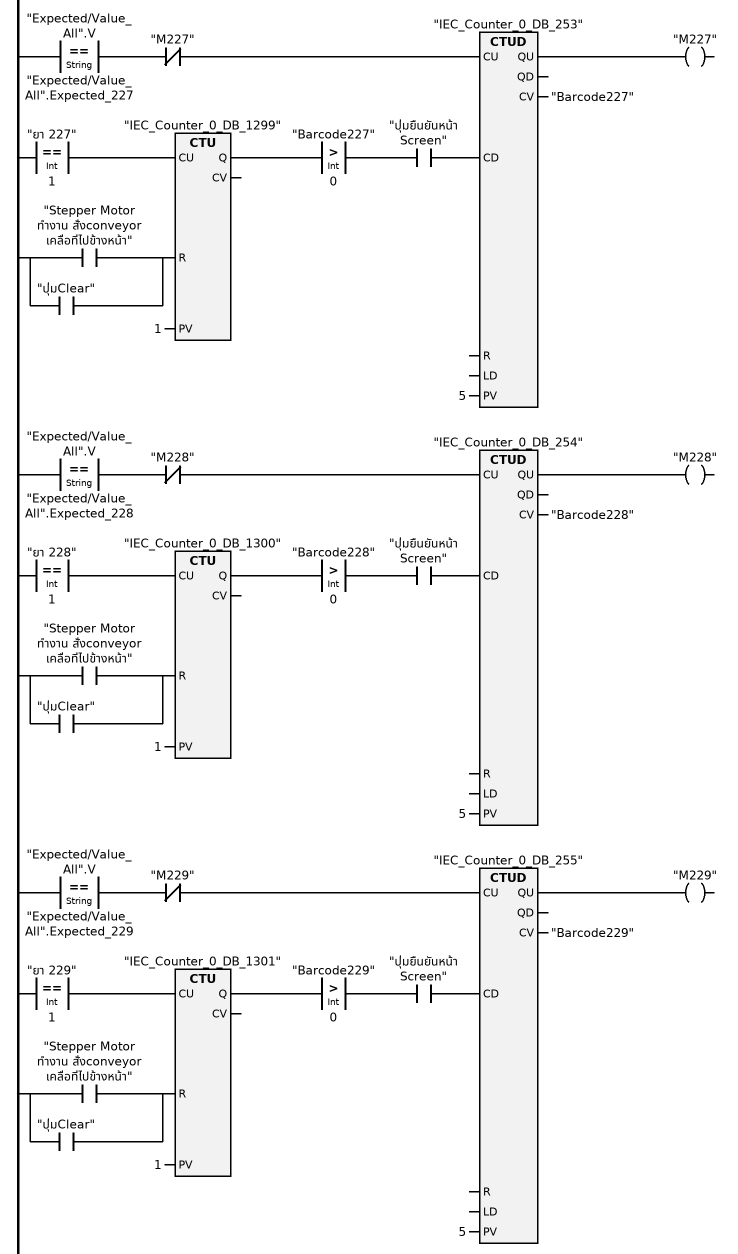
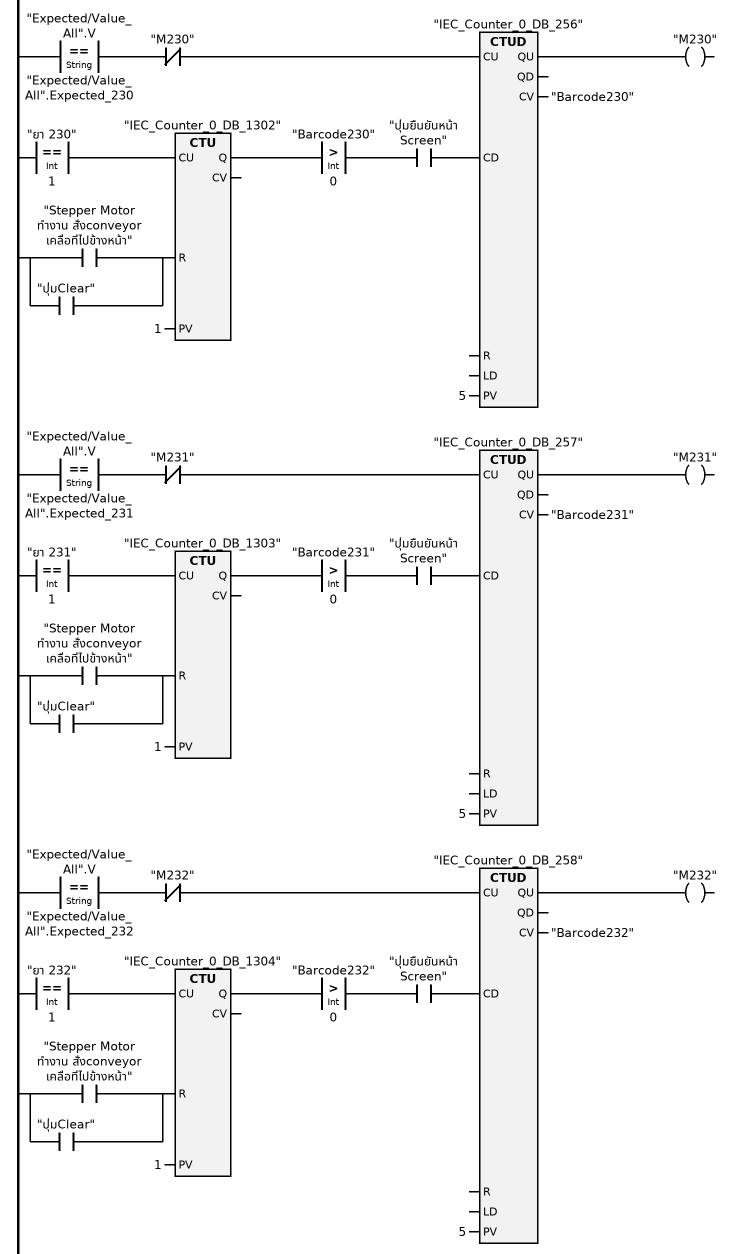
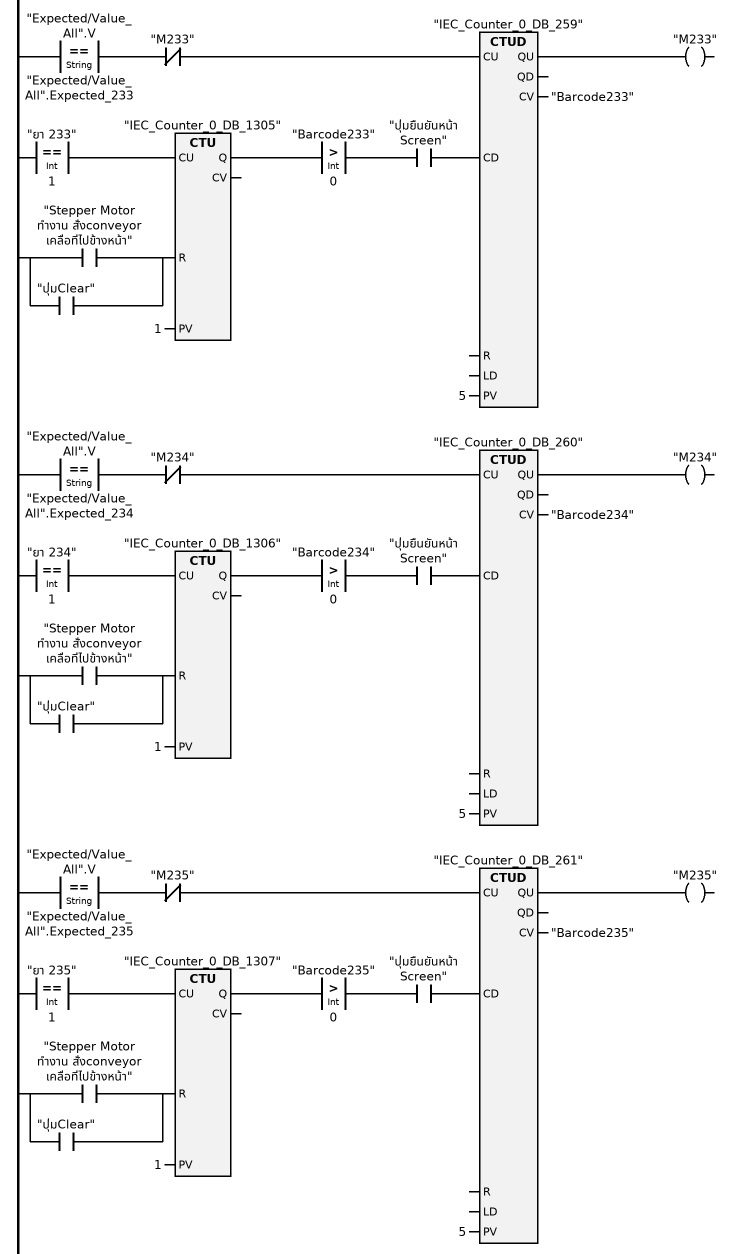
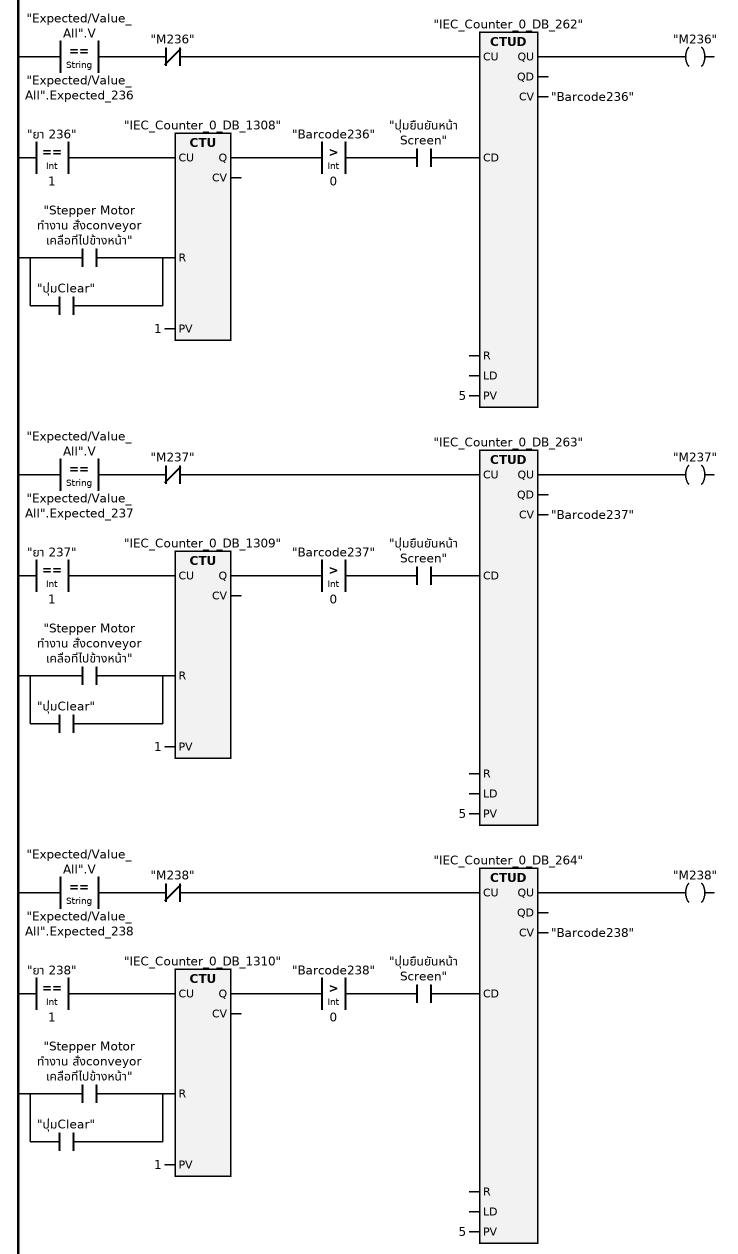
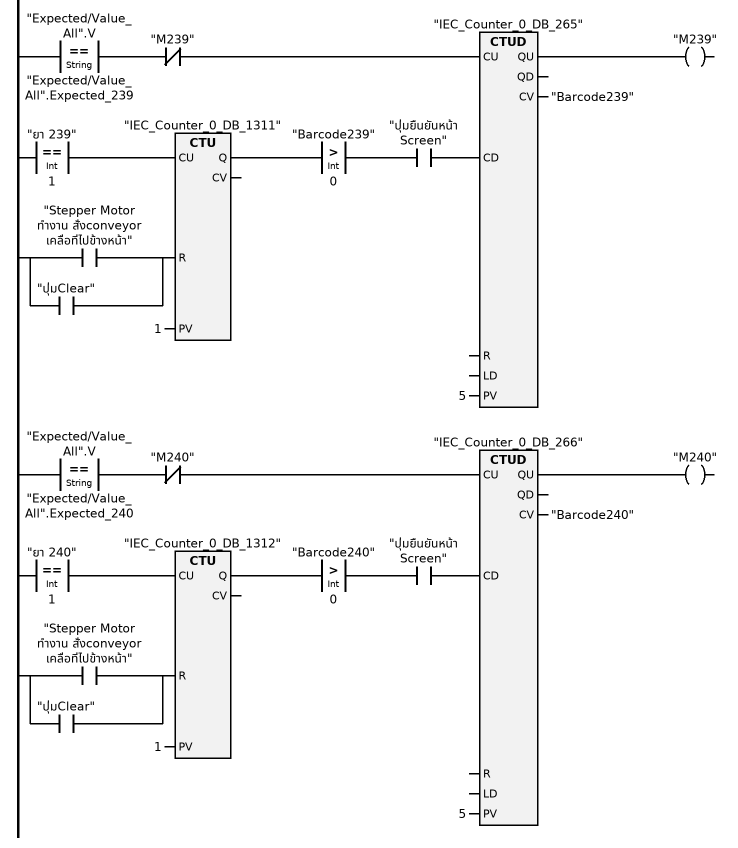
   "IEC_Counter_0_DB_1293".CTU(CU := "ยา 221" = 1,
                           R := "Stepper Motor ทำงาน สั่งconveyor เคลื่อที่ไปข้างหน้า" OR "ปุ่มClear",
                           PV := 1);
   "IEC_Counter_0_DB_247".CTUD(CU := ("Expected/Value_All".V = "Expected/Value_All".Expected_221) AND NOT "M221",
                           CD := "IEC_Counter_0_DB_1293".Q AND ("Barcode221" > 0) AND "ปุ่มยืนยันหน้า Screen",
                           PV := 5,
                           CV => "Barcode221");
   "M221" := "IEC_Counter_0_DB_247".QU;
   "IEC_Counter_0_DB_1294".CTU(CU := "ยา 222" = 1,
                           R := "Stepper Motor ทำงาน สั่งconveyor เคลื่อที่ไปข้างหน้า" OR "ปุ่มClear",
                           PV := 1);
   "IEC_Counter_0_DB_248".CTUD(CU := ("Expected/Value_All".V = "Expected/Value_All".Expected_222) AND NOT "M222",
                           CD := "IEC_Counter_0_DB_1294".Q AND ("Barcode222" > 0) AND "ปุ่มยืนยันหน้า Screen",
                           PV := 5,
                           CV => "Barcode222");
   "M222" := "IEC_Counter_0_DB_248".QU;
   "IEC_Counter_0_DB_1295".CTU(CU := "ยา 223" = 1,
                           R := "Stepper Motor ทำงาน สั่งconveyor เคลื่อที่ไปข้างหน้า" OR "ปุ่มClear",
                           PV := 1);
   "IEC_Counter_0_DB_249".CTUD(CU := ("Expected/Value_All".V = "Expected/Value_All".Expected_223) AND NOT "M223",
                           CD := "IEC_Counter_0_DB_1295".Q AND ("Barcode223" > 0) AND "ปุ่มยืนยันหน้า Screen",
                           PV := 5,
                           CV => "Barcode223");
   "M223" := "IEC_Counter_0_DB_249".QU;
   "IEC_Counter_0_DB_1296".CTU(CU := "ยา 224" = 1,
                           R := "Stepper Motor ทำงาน สั่งconveyor เคลื่อที่ไปข้างหน้า" OR "ปุ่มClear",
                           PV := 1);
   "IEC_Counter_0_DB_250".CTUD(CU := ("Expected/Value_All".V = "Expected/Value_All".Expected_224) AND NOT "M224",
                           CD := "IEC_Counter_0_DB_1296".Q AND ("Barcode224" > 0) AND "ปุ่มยืนยันหน้า Screen",
                           PV := 5,
                           CV => "Barcode224");
   "M224" := "IEC_Counter_0_DB_250".QU;
   "IEC_Counter_0_DB_1297".CTU(CU := "ยา 225" = 1,
                           R := "Stepper Motor ทำงาน สั่งconveyor เคลื่อที่ไปข้างหน้า" OR "ปุ่มClear",
                           PV := 1);
   "IEC_Counter_0_DB_251".CTUD(CU := ("Expected/Value_All".V = "Expected/Value_All".Expected_225) AND NOT "M225",
                           CD := "IEC_Counter_0_DB_1297".Q AND ("Barcode225" > 0) AND "ปุ่มยืนยันหน้า Screen",
                           PV := 5,
                           CV => "Barcode225");
   "M225" := "IEC_Counter_0_DB_251".QU;
   "IEC_Counter_0_DB_1298".CTU(CU := "ยา 226" = 1,
                           R := "Stepper Motor ทำงาน สั่งconveyor เคลื่อที่ไปข้างหน้า" OR "ปุ่มClear",
                           PV := 1);
   "IEC_Counter_0_DB_252".CTUD(CU := ("Expected/Value_All".V = "Expected/Value_All".Expected_226) AND NOT "M226",
                           CD := "IEC_Counter_0_DB_1298".Q AND ("Barcode226" > 0) AND "ปุ่มยืนยันหน้า Screen",
                           PV := 5,
                           CV => "Barcode226");
   "M226" := "IEC_Counter_0_DB_252".QU;
   "IEC_Counter_0_DB_1299".CTU(CU := "ยา 227" = 1,
                           R := "Stepper Motor ทำงาน สั่งconveyor เคลื่อที่ไปข้างหน้า" OR "ปุ่มClear",
                           PV := 1);
   "IEC_Counter_0_DB_253".CTUD(CU := ("Expected/Value_All".V = "Expected/Value_All".Expected_227) AND NOT "M227",
                           CD := "IEC_Counter_0_DB_1299".Q AND ("Barcode227" > 0) AND "ปุ่มยืนยันหน้า Screen",
                           PV := 5,
                           CV => "Barcode227");
   "M227" := "IEC_Counter_0_DB_253".QU;
   "IEC_Counter_0_DB_1300".CTU(CU := "ยา 228" = 1,
                           R := "Stepper Motor ทำงาน สั่งconveyor เคลื่อที่ไปข้างหน้า" OR "ปุ่มClear",
                           PV := 1);
   "IEC_Counter_0_DB_254".CTUD(CU := ("Expected/Value_All".V = "Expected/Value_All".Expected_228) AND NOT "M228",
                           CD := "IEC_Counter_0_DB_1300".Q AND ("Barcode228" > 0) AND "ปุ่มยืนยันหน้า Screen",
                           PV := 5,
                           CV => "Barcode228");
   "M228" := "IEC_Counter_0_DB_254".QU;
   "IEC_Counter_0_DB_1301".CTU(CU := "ยา 229" = 1,
                           R := "Stepper Motor ทำงาน สั่งconveyor เคลื่อที่ไปข้างหน้า" OR "ปุ่มClear",
                           PV := 1);
   "IEC_Counter_0_DB_255".CTUD(CU := ("Expected/Value_All".V = "Expected/Value_All".Expected_229) AND NOT "M229",
                           CD := "IEC_Counter_0_DB_1301".Q AND ("Barcode229" > 0) AND "ปุ่มยืนยันหน้า Screen",
                           PV := 5,
                           CV => "Barcode229");
   "M229" := "IEC_Counter_0_DB_255".QU;
   "IEC_Counter_0_DB_1302".CTU(CU := "ยา 230" = 1,
                           R := "Stepper Motor ทำงาน สั่งconveyor เคลื่อที่ไปข้างหน้า" OR "ปุ่มClear",
                           PV := 1);
   "IEC_Counter_0_DB_256".CTUD(CU := ("Expected/Value_All".V = "Expected/Value_All".Expected_230) AND NOT "M230",
                           CD := "IEC_Counter_0_DB_1302".Q AND ("Barcode230" > 0) AND "ปุ่มยืนยันหน้า Screen",
                           PV := 5,
                           CV => "Barcode230");
   "M230" := "IEC_Counter_0_DB_256".QU;
   "IEC_Counter_0_DB_1303".CTU(CU := "ยา 231" = 1,
                           R := "Stepper Motor ทำงาน สั่งconveyor เคลื่อที่ไปข้างหน้า" OR "ปุ่มClear",
                           PV := 1);
   "IEC_Counter_0_DB_257".CTUD(CU := ("Expected/Value_All".V = "Expected/Value_All".Expected_231) AND NOT "M231",
                           CD := "IEC_Counter_0_DB_1303".Q AND ("Barcode231" > 0) AND "ปุ่มยืนยันหน้า Screen",
                           PV := 5,
                           CV => "Barcode231");
   "M231" := "IEC_Counter_0_DB_257".QU;
   "IEC_Counter_0_DB_1304".CTU(CU := "ยา 232" = 1,
                           R := "Stepper Motor ทำงาน สั่งconveyor เคลื่อที่ไปข้างหน้า" OR "ปุ่มClear",
                           PV := 1);
   "IEC_Counter_0_DB_258".CTUD(CU := ("Expected/Value_All".V = "Expected/Value_All".Expected_232) AND NOT "M232",
                           CD := "IEC_Counter_0_DB_1304".Q AND ("Barcode232" > 0) AND "ปุ่มยืนยันหน้า Screen",
                           PV := 5,
                           CV => "Barcode232");
   "M232" := "IEC_Counter_0_DB_258".QU;
   "IEC_Counter_0_DB_1305".CTU(CU := "ยา 233" = 1,
                           R := "Stepper Motor ทำงาน สั่งconveyor เคลื่อที่ไปข้างหน้า" OR "ปุ่มClear",
                           PV := 1);
   "IEC_Counter_0_DB_259".CTUD(CU := ("Expected/Value_All".V = "Expected/Value_All".Expected_233) AND NOT "M233",
                           CD := "IEC_Counter_0_DB_1305".Q AND ("Barcode233" > 0) AND "ปุ่มยืนยันหน้า Screen",
                           PV := 5,
                           CV => "Barcode233");
   "M233" := "IEC_Counter_0_DB_259".QU;
   "IEC_Counter_0_DB_1306".CTU(CU := "ยา 234" = 1,
                           R := "Stepper Motor ทำงาน สั่งconveyor เคลื่อที่ไปข้างหน้า" OR "ปุ่มClear",
                           PV := 1);
   "IEC_Counter_0_DB_260".CTUD(CU := ("Expected/Value_All".V = "Expected/Value_All".Expected_234) AND NOT "M234",
                           CD := "IEC_Counter_0_DB_1306".Q AND ("Barcode234" > 0) AND "ปุ่มยืนยันหน้า Screen",
                           PV := 5,
                           CV => "Barcode234");
   "M234" := "IEC_Counter_0_DB_260".QU;
   "IEC_Counter_0_DB_1307".CTU(CU := "ยา 235" = 1,
                           R := "Stepper Motor ทำงาน สั่งconveyor เคลื่อที่ไปข้างหน้า" OR "ปุ่มClear",
                           PV := 1);
   "IEC_Counter_0_DB_261".CTUD(CU := ("Expected/Value_All".V = "Expected/Value_All".Expected_235) AND NOT "M235",
                           CD := "IEC_Counter_0_DB_1307".Q AND ("Barcode235" > 0) AND "ปุ่มยืนยันหน้า Screen",
                           PV := 5,
                           CV => "Barcode235");
   "M235" := "IEC_Counter_0_DB_261".QU;
   "IEC_Counter_0_DB_1308".CTU(CU := "ยา 236" = 1,
                           R := "Stepper Motor ทำงาน สั่งconveyor เคลื่อที่ไปข้างหน้า" OR "ปุ่มClear",
                           PV := 1);
   "IEC_Counter_0_DB_262".CTUD(CU := ("Expected/Value_All".V = "Expected/Value_All".Expected_236) AND NOT "M236",
                           CD := "IEC_Counter_0_DB_1308".Q AND ("Barcode236" > 0) AND "ปุ่มยืนยันหน้า Screen",
                           PV := 5,
                           CV => "Barcode236");
   "M236" := "IEC_Counter_0_DB_262".QU;
   "IEC_Counter_0_DB_1309".CTU(CU := "ยา 237" = 1,
                           R := "Stepper Motor ทำงาน สั่งconveyor เคลื่อที่ไปข้างหน้า" OR "ปุ่มClear",
                           PV := 1);
   "IEC_Counter_0_DB_263".CTUD(CU := ("Expected/Value_All".V = "Expected/Value_All".Expected_237) AND NOT "M237",
                           CD := "IEC_Counter_0_DB_1309".Q AND ("Barcode237" > 0) AND "ปุ่มยืนยันหน้า Screen",
                           PV := 5,
                           CV => "Barcode237");
   "M237" := "IEC_Counter_0_DB_263".QU;
   "IEC_Counter_0_DB_1310".CTU(CU := "ยา 238" = 1,
                           R := "Stepper Motor ทำงาน สั่งconveyor เคลื่อที่ไปข้างหน้า" OR "ปุ่มClear",
                           PV := 1);
   "IEC_Counter_0_DB_264".CTUD(CU := ("Expected/Value_All".V = "Expected/Value_All".Expected_238) AND NOT "M238",
                           CD := "IEC_Counter_0_DB_1310".Q AND ("Barcode238" > 0) AND "ปุ่มยืนยันหน้า Screen",
                           PV := 5,
                           CV => "Barcode238");
   "M238" := "IEC_Counter_0_DB_264".QU;
   "IEC_Counter_0_DB_1311".CTU(CU := "ยา 239" = 1,
                           R := "Stepper Motor ทำงาน สั่งconveyor เคลื่อที่ไปข้างหน้า" OR "ปุ่มClear",
                           PV := 1);
   "IEC_Counter_0_DB_265".CTUD(CU := ("Expected/Value_All".V = "Expected/Value_All".Expected_239) AND NOT "M239",
                           CD := "IEC_Counter_0_DB_1311".Q AND ("Barcode239" > 0) AND "ปุ่มยืนยันหน้า Screen",
                           PV := 5,
                           CV => "Barcode239");
   "M239" := "IEC_Counter_0_DB_265".QU;
   "IEC_Counter_0_DB_1312".CTU(CU := "ยา 240" = 1,
                           R := "Stepper Motor ทำงาน สั่งconveyor เคลื่อที่ไปข้างหน้า" OR "ปุ่มClear",
                           PV := 1);
   "IEC_Counter_0_DB_266".CTUD(CU := ("Expected/Value_All".V = "Expected/Value_All".Expected_240) AND NOT "M240",
                           CD := "IEC_Counter_0_DB_1312".Q AND ("Barcode240" > 0) AND "ปุ่มยืนยันหน้า Screen",
                           PV := 5,
                           CV => "Barcode240");
   "M240" := "IEC_Counter_0_DB_266".QU;
END_REGION

REGION Network 13
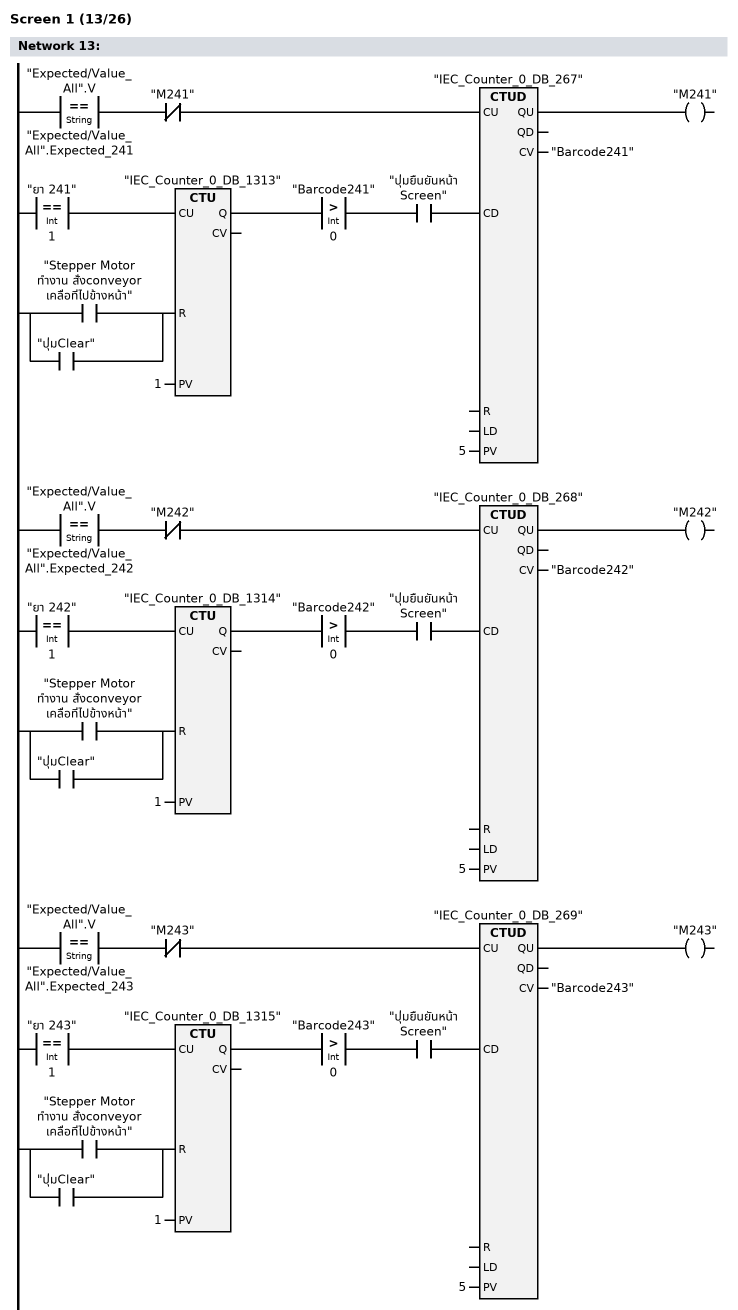
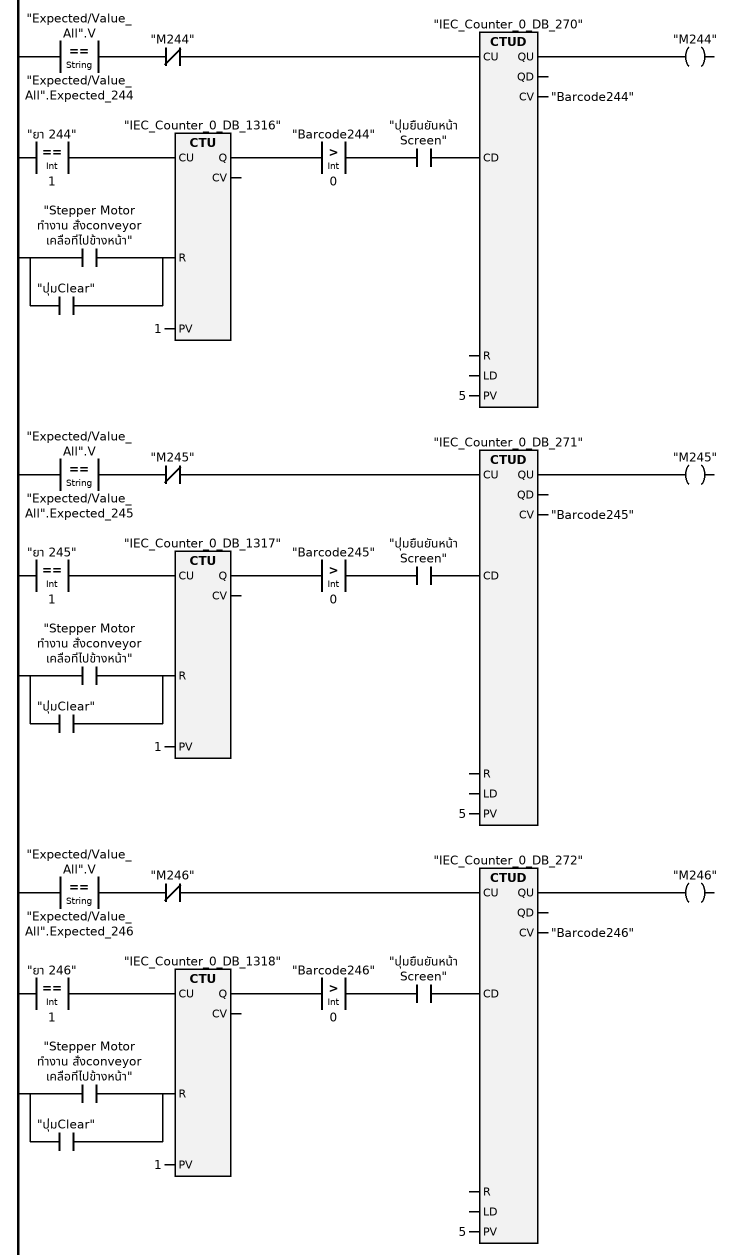
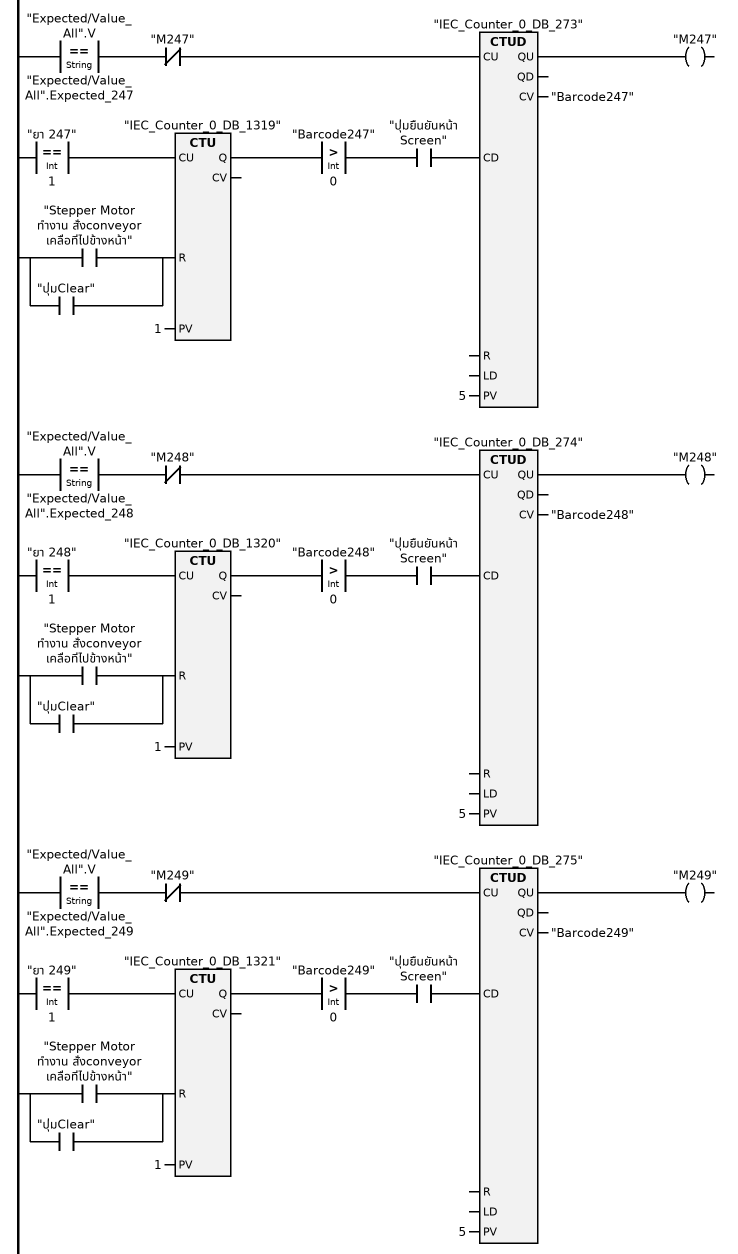
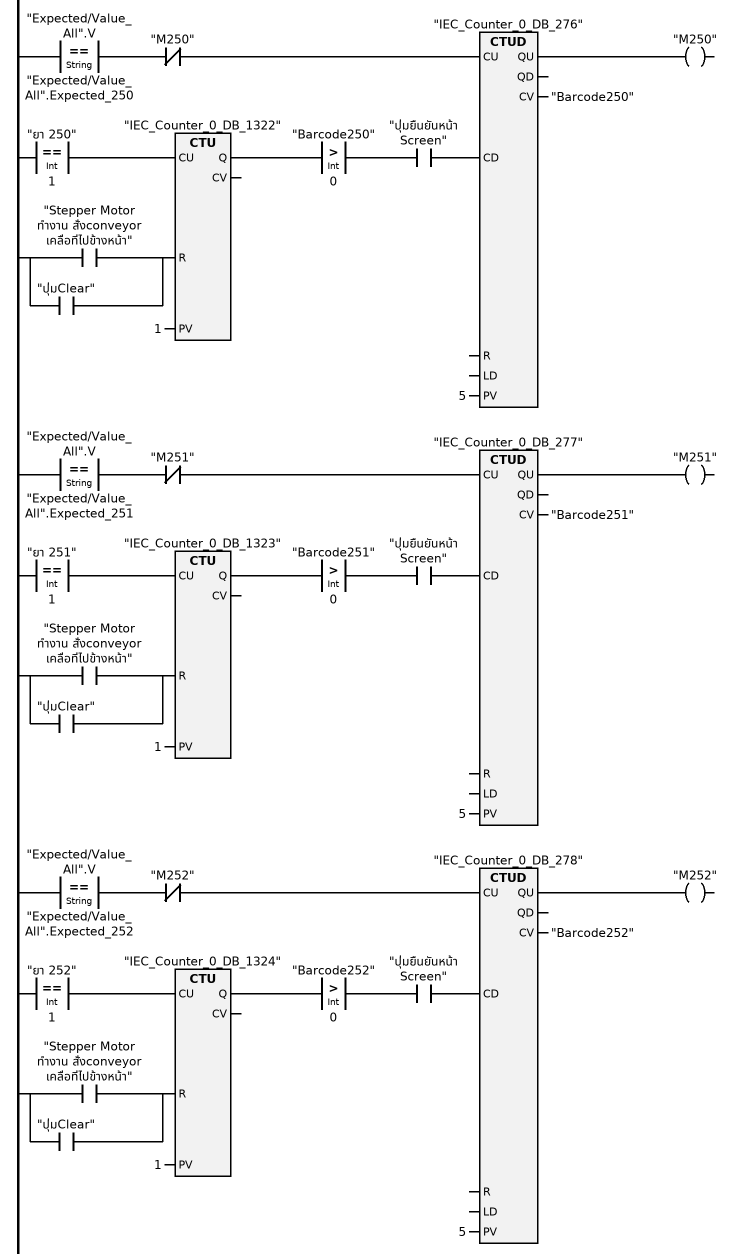
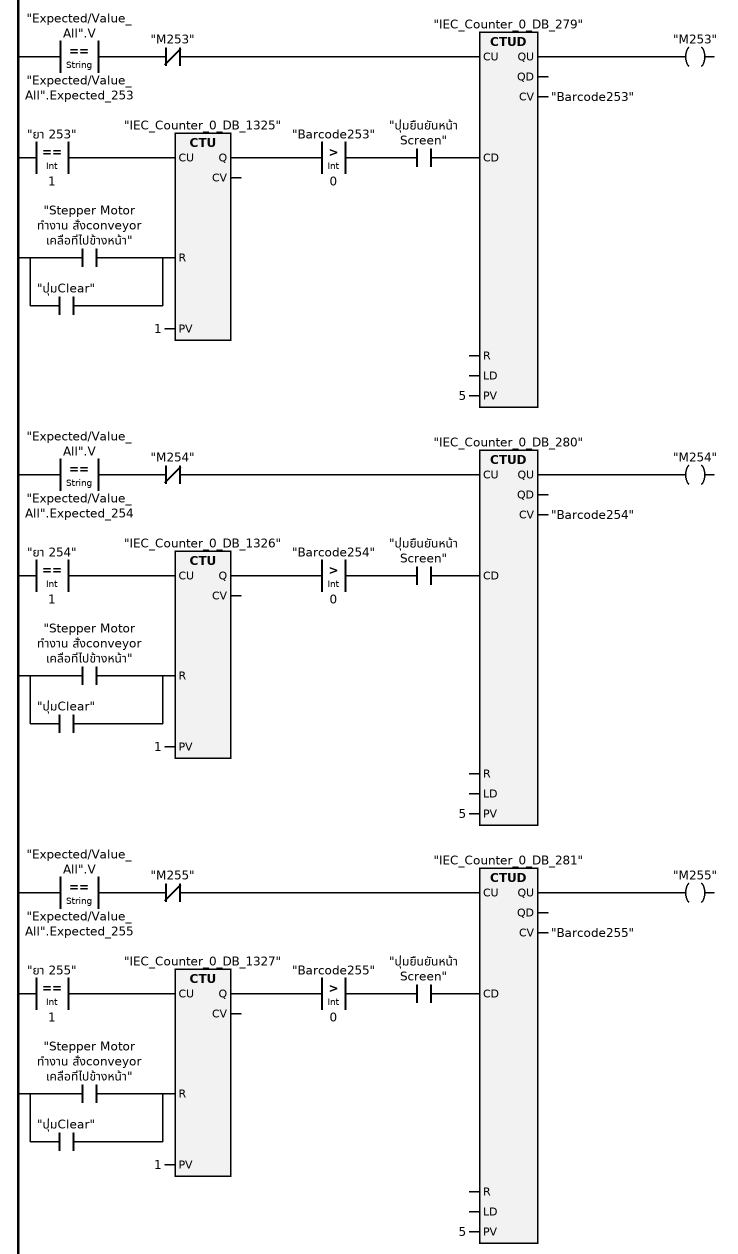
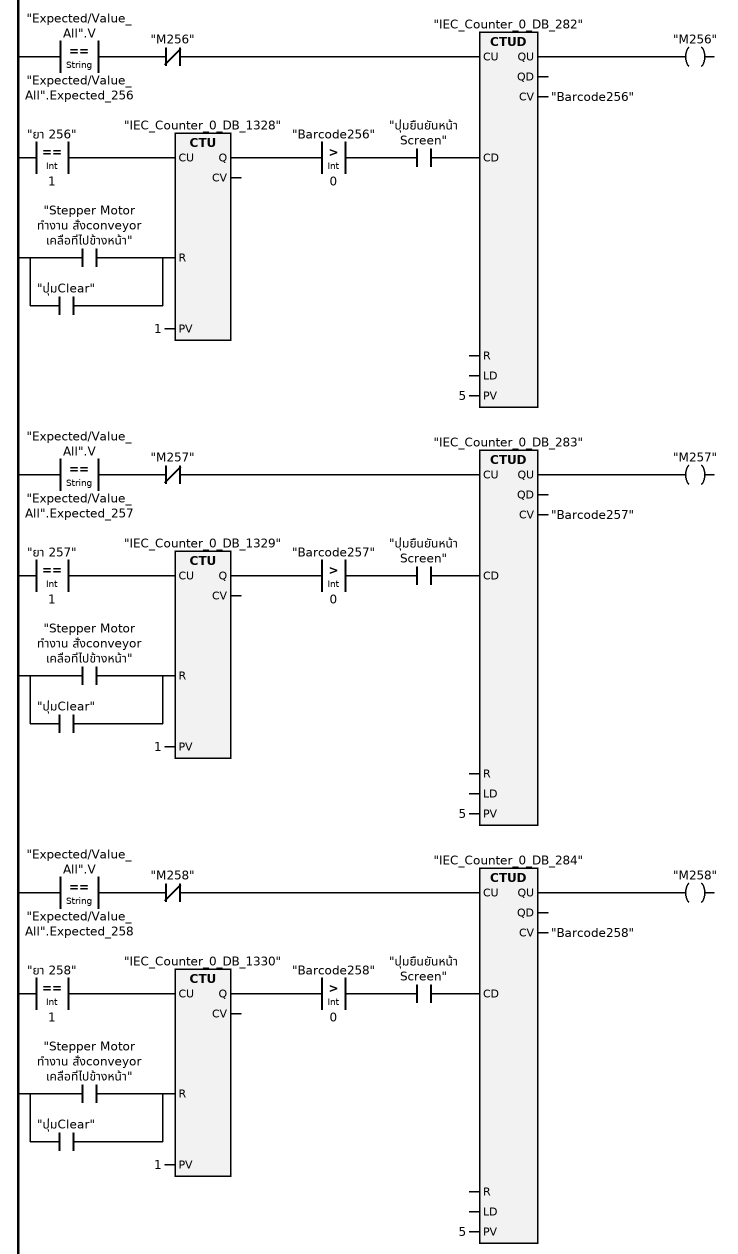
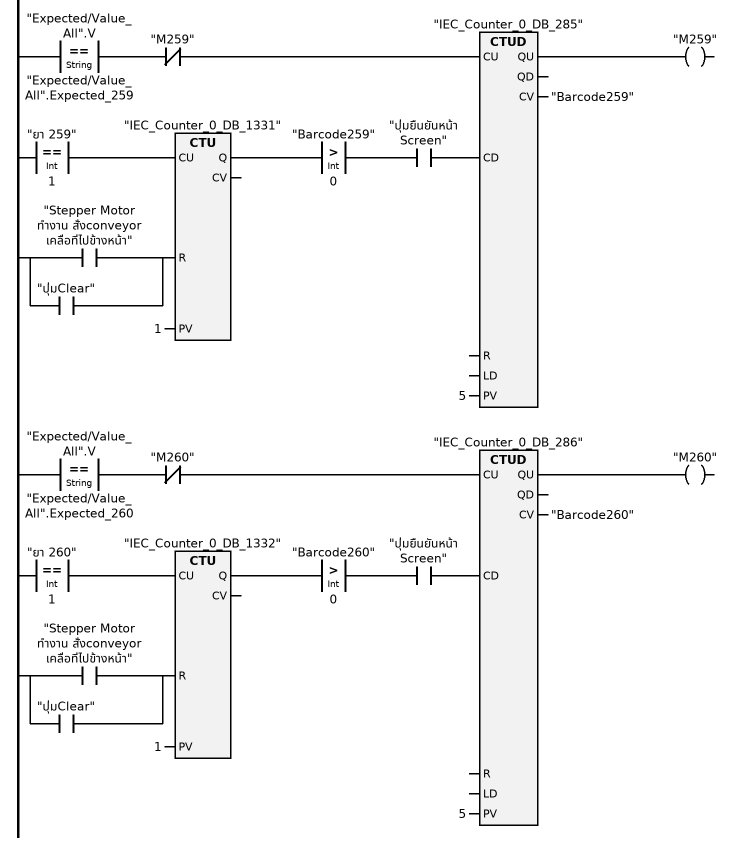
   "IEC_Counter_0_DB_1313".CTU(CU := "ยา 241" = 1,
                           R := "Stepper Motor ทำงาน สั่งconveyor เคลื่อที่ไปข้างหน้า" OR "ปุ่มClear",
                           PV := 1);
   "IEC_Counter_0_DB_267".CTUD(CU := ("Expected/Value_All".V = "Expected/Value_All".Expected_241) AND NOT "M241",
                           CD := "IEC_Counter_0_DB_1313".Q AND ("Barcode241" > 0) AND "ปุ่มยืนยันหน้า Screen",
                           PV := 5,
                           CV => "Barcode241");
   "M241" := "IEC_Counter_0_DB_267".QU;
   "IEC_Counter_0_DB_1314".CTU(CU := "ยา 242" = 1,
                           R := "Stepper Motor ทำงาน สั่งconveyor เคลื่อที่ไปข้างหน้า" OR "ปุ่มClear",
                           PV := 1);
   "IEC_Counter_0_DB_268".CTUD(CU := ("Expected/Value_All".V = "Expected/Value_All".Expected_242) AND NOT "M242",
                           CD := "IEC_Counter_0_DB_1314".Q AND ("Barcode242" > 0) AND "ปุ่มยืนยันหน้า Screen",
                           PV := 5,
                           CV => "Barcode242");
   "M242" := "IEC_Counter_0_DB_268".QU;
   "IEC_Counter_0_DB_1315".CTU(CU := "ยา 243" = 1,
                           R := "Stepper Motor ทำงาน สั่งconveyor เคลื่อที่ไปข้างหน้า" OR "ปุ่มClear",
                           PV := 1);
   "IEC_Counter_0_DB_269".CTUD(CU := ("Expected/Value_All".V = "Expected/Value_All".Expected_243) AND NOT "M243",
                           CD := "IEC_Counter_0_DB_1315".Q AND ("Barcode243" > 0) AND "ปุ่มยืนยันหน้า Screen",
                           PV := 5,
                           CV => "Barcode243");
   "M243" := "IEC_Counter_0_DB_269".QU;
   "IEC_Counter_0_DB_1316".CTU(CU := "ยา 244" = 1,
                           R := "Stepper Motor ทำงาน สั่งconveyor เคลื่อที่ไปข้างหน้า" OR "ปุ่มClear",
                           PV := 1);
   "IEC_Counter_0_DB_270".CTUD(CU := ("Expected/Value_All".V = "Expected/Value_All".Expected_244) AND NOT "M244",
                           CD := "IEC_Counter_0_DB_1316".Q AND ("Barcode244" > 0) AND "ปุ่มยืนยันหน้า Screen",
                           PV := 5,
                           CV => "Barcode244");
   "M244" := "IEC_Counter_0_DB_270".QU;
   "IEC_Counter_0_DB_1317".CTU(CU := "ยา 245" = 1,
                           R := "Stepper Motor ทำงาน สั่งconveyor เคลื่อที่ไปข้างหน้า" OR "ปุ่มClear",
                           PV := 1);
   "IEC_Counter_0_DB_271".CTUD(CU := ("Expected/Value_All".V = "Expected/Value_All".Expected_245) AND NOT "M245",
                           CD := "IEC_Counter_0_DB_1317".Q AND ("Barcode245" > 0) AND "ปุ่มยืนยันหน้า Screen",
                           PV := 5,
                           CV => "Barcode245");
   "M245" := "IEC_Counter_0_DB_271".QU;
   "IEC_Counter_0_DB_1318".CTU(CU := "ยา 246" = 1,
                           R := "Stepper Motor ทำงาน สั่งconveyor เคลื่อที่ไปข้างหน้า" OR "ปุ่มClear",
                           PV := 1);
   "IEC_Counter_0_DB_272".CTUD(CU := ("Expected/Value_All".V = "Expected/Value_All".Expected_246) AND NOT "M246",
                           CD := "IEC_Counter_0_DB_1318".Q AND ("Barcode246" > 0) AND "ปุ่มยืนยันหน้า Screen",
                           PV := 5,
                           CV => "Barcode246");
   "M246" := "IEC_Counter_0_DB_272".QU;
   "IEC_Counter_0_DB_1319".CTU(CU := "ยา 247" = 1,
                           R := "Stepper Motor ทำงาน สั่งconveyor เคลื่อที่ไปข้างหน้า" OR "ปุ่มClear",
                           PV := 1);
   "IEC_Counter_0_DB_273".CTUD(CU := ("Expected/Value_All".V = "Expected/Value_All".Expected_247) AND NOT "M247",
                           CD := "IEC_Counter_0_DB_1319".Q AND ("Barcode247" > 0) AND "ปุ่มยืนยันหน้า Screen",
                           PV := 5,
                           CV => "Barcode247");
   "M247" := "IEC_Counter_0_DB_273".QU;
   "IEC_Counter_0_DB_1320".CTU(CU := "ยา 248" = 1,
                           R := "Stepper Motor ทำงาน สั่งconveyor เคลื่อที่ไปข้างหน้า" OR "ปุ่มClear",
                           PV := 1);
   "IEC_Counter_0_DB_274".CTUD(CU := ("Expected/Value_All".V = "Expected/Value_All".Expected_248) AND NOT "M248",
                           CD := "IEC_Counter_0_DB_1320".Q AND ("Barcode248" > 0) AND "ปุ่มยืนยันหน้า Screen",
                           PV := 5,
                           CV => "Barcode248");
   "M248" := "IEC_Counter_0_DB_274".QU;
   "IEC_Counter_0_DB_1321".CTU(CU := "ยา 249" = 1,
                           R := "Stepper Motor ทำงาน สั่งconveyor เคลื่อที่ไปข้างหน้า" OR "ปุ่มClear",
                           PV := 1);
   "IEC_Counter_0_DB_275".CTUD(CU := ("Expected/Value_All".V = "Expected/Value_All".Expected_249) AND NOT "M249",
                           CD := "IEC_Counter_0_DB_1321".Q AND ("Barcode249" > 0) AND "ปุ่มยืนยันหน้า Screen",
                           PV := 5,
                           CV => "Barcode249");
   "M249" := "IEC_Counter_0_DB_275".QU;
   "IEC_Counter_0_DB_1322".CTU(CU := "ยา 250" = 1,
                           R := "Stepper Motor ทำงาน สั่งconveyor เคลื่อที่ไปข้างหน้า" OR "ปุ่มClear",
                           PV := 1);
   "IEC_Counter_0_DB_276".CTUD(CU := ("Expected/Value_All".V = "Expected/Value_All".Expected_250) AND NOT "M250",
                           CD := "IEC_Counter_0_DB_1322".Q AND ("Barcode250" > 0) AND "ปุ่มยืนยันหน้า Screen",
                           PV := 5,
                           CV => "Barcode250");
   "M250" := "IEC_Counter_0_DB_276".QU;
   "IEC_Counter_0_DB_1323".CTU(CU := "ยา 251" = 1,
                           R := "Stepper Motor ทำงาน สั่งconveyor เคลื่อที่ไปข้างหน้า" OR "ปุ่มClear",
                           PV := 1);
   "IEC_Counter_0_DB_277".CTUD(CU := ("Expected/Value_All".V = "Expected/Value_All".Expected_251) AND NOT "M251",
                           CD := "IEC_Counter_0_DB_1323".Q AND ("Barcode251" > 0) AND "ปุ่มยืนยันหน้า Screen",
                           PV := 5,
                           CV => "Barcode251");
   "M251" := "IEC_Counter_0_DB_277".QU;
   "IEC_Counter_0_DB_1324".CTU(CU := "ยา 252" = 1,
                           R := "Stepper Motor ทำงาน สั่งconveyor เคลื่อที่ไปข้างหน้า" OR "ปุ่มClear",
                           PV := 1);
   "IEC_Counter_0_DB_278".CTUD(CU := ("Expected/Value_All".V = "Expected/Value_All".Expected_252) AND NOT "M252",
                           CD := "IEC_Counter_0_DB_1324".Q AND ("Barcode252" > 0) AND "ปุ่มยืนยันหน้า Screen",
                           PV := 5,
                           CV => "Barcode252");
   "M252" := "IEC_Counter_0_DB_278".QU;
   "IEC_Counter_0_DB_1325".CTU(CU := "ยา 253" = 1,
                           R := "Stepper Motor ทำงาน สั่งconveyor เคลื่อที่ไปข้างหน้า" OR "ปุ่มClear",
                           PV := 1);
   "IEC_Counter_0_DB_279".CTUD(CU := ("Expected/Value_All".V = "Expected/Value_All".Expected_253) AND NOT "M253",
                           CD := "IEC_Counter_0_DB_1325".Q AND ("Barcode253" > 0) AND "ปุ่มยืนยันหน้า Screen",
                           PV := 5,
                           CV => "Barcode253");
   "M253" := "IEC_Counter_0_DB_279".QU;
   "IEC_Counter_0_DB_1326".CTU(CU := "ยา 254" = 1,
                           R := "Stepper Motor ทำงาน สั่งconveyor เคลื่อที่ไปข้างหน้า" OR "ปุ่มClear",
                           PV := 1);
   "IEC_Counter_0_DB_280".CTUD(CU := ("Expected/Value_All".V = "Expected/Value_All".Expected_254) AND NOT "M254",
                           CD := "IEC_Counter_0_DB_1326".Q AND ("Barcode254" > 0) AND "ปุ่มยืนยันหน้า Screen",
                           PV := 5,
                           CV => "Barcode254");
   "M254" := "IEC_Counter_0_DB_280".QU;
   "IEC_Counter_0_DB_1327".CTU(CU := "ยา 255" = 1,
                           R := "Stepper Motor ทำงาน สั่งconveyor เคลื่อที่ไปข้างหน้า" OR "ปุ่มClear",
                           PV := 1);
   "IEC_Counter_0_DB_281".CTUD(CU := ("Expected/Value_All".V = "Expected/Value_All".Expected_255) AND NOT "M255",
                           CD := "IEC_Counter_0_DB_1327".Q AND ("Barcode255" > 0) AND "ปุ่มยืนยันหน้า Screen",
                           PV := 5,
                           CV => "Barcode255");
   "M255" := "IEC_Counter_0_DB_281".QU;
   "IEC_Counter_0_DB_1328".CTU(CU := "ยา 256" = 1,
                           R := "Stepper Motor ทำงาน สั่งconveyor เคลื่อที่ไปข้างหน้า" OR "ปุ่มClear",
                           PV := 1);
   "IEC_Counter_0_DB_282".CTUD(CU := ("Expected/Value_All".V = "Expected/Value_All".Expected_256) AND NOT "M256",
                           CD := "IEC_Counter_0_DB_1328".Q AND ("Barcode256" > 0) AND "ปุ่มยืนยันหน้า Screen",
                           PV := 5,
                           CV => "Barcode256");
   "M256" := "IEC_Counter_0_DB_282".QU;
   "IEC_Counter_0_DB_1329".CTU(CU := "ยา 257" = 1,
                           R := "Stepper Motor ทำงาน สั่งconveyor เคลื่อที่ไปข้างหน้า" OR "ปุ่มClear",
                           PV := 1);
   "IEC_Counter_0_DB_283".CTUD(CU := ("Expected/Value_All".V = "Expected/Value_All".Expected_257) AND NOT "M257",
                           CD := "IEC_Counter_0_DB_1329".Q AND ("Barcode257" > 0) AND "ปุ่มยืนยันหน้า Screen",
                           PV := 5,
                           CV => "Barcode257");
   "M257" := "IEC_Counter_0_DB_283".QU;
   "IEC_Counter_0_DB_1330".CTU(CU := "ยา 258" = 1,
                           R := "Stepper Motor ทำงาน สั่งconveyor เคลื่อที่ไปข้างหน้า" OR "ปุ่มClear",
                           PV := 1);
   "IEC_Counter_0_DB_284".CTUD(CU := ("Expected/Value_All".V = "Expected/Value_All".Expected_258) AND NOT "M258",
                           CD := "IEC_Counter_0_DB_1330".Q AND ("Barcode258" > 0) AND "ปุ่มยืนยันหน้า Screen",
                           PV := 5,
                           CV => "Barcode258");
   "M258" := "IEC_Counter_0_DB_284".QU;
   "IEC_Counter_0_DB_1331".CTU(CU := "ยา 259" = 1,
                           R := "Stepper Motor ทำงาน สั่งconveyor เคลื่อที่ไปข้างหน้า" OR "ปุ่มClear",
                           PV := 1);
   "IEC_Counter_0_DB_285".CTUD(CU := ("Expected/Value_All".V = "Expected/Value_All".Expected_259) AND NOT "M259",
                           CD := "IEC_Counter_0_DB_1331".Q AND ("Barcode259" > 0) AND "ปุ่มยืนยันหน้า Screen",
                           PV := 5,
                           CV => "Barcode259");
   "M259" := "IEC_Counter_0_DB_285".QU;
   "IEC_Counter_0_DB_1332".CTU(CU := "ยา 260" = 1,
                           R := "Stepper Motor ทำงาน สั่งconveyor เคลื่อที่ไปข้างหน้า" OR "ปุ่มClear",
                           PV := 1);
   "IEC_Counter_0_DB_286".CTUD(CU := ("Expected/Value_All".V = "Expected/Value_All".Expected_260) AND NOT "M260",
                           CD := "IEC_Counter_0_DB_1332".Q AND ("Barcode260" > 0) AND "ปุ่มยืนยันหน้า Screen",
                           PV := 5,
                           CV => "Barcode260");
   "M260" := "IEC_Counter_0_DB_286".QU;
END_REGION

REGION Network 14
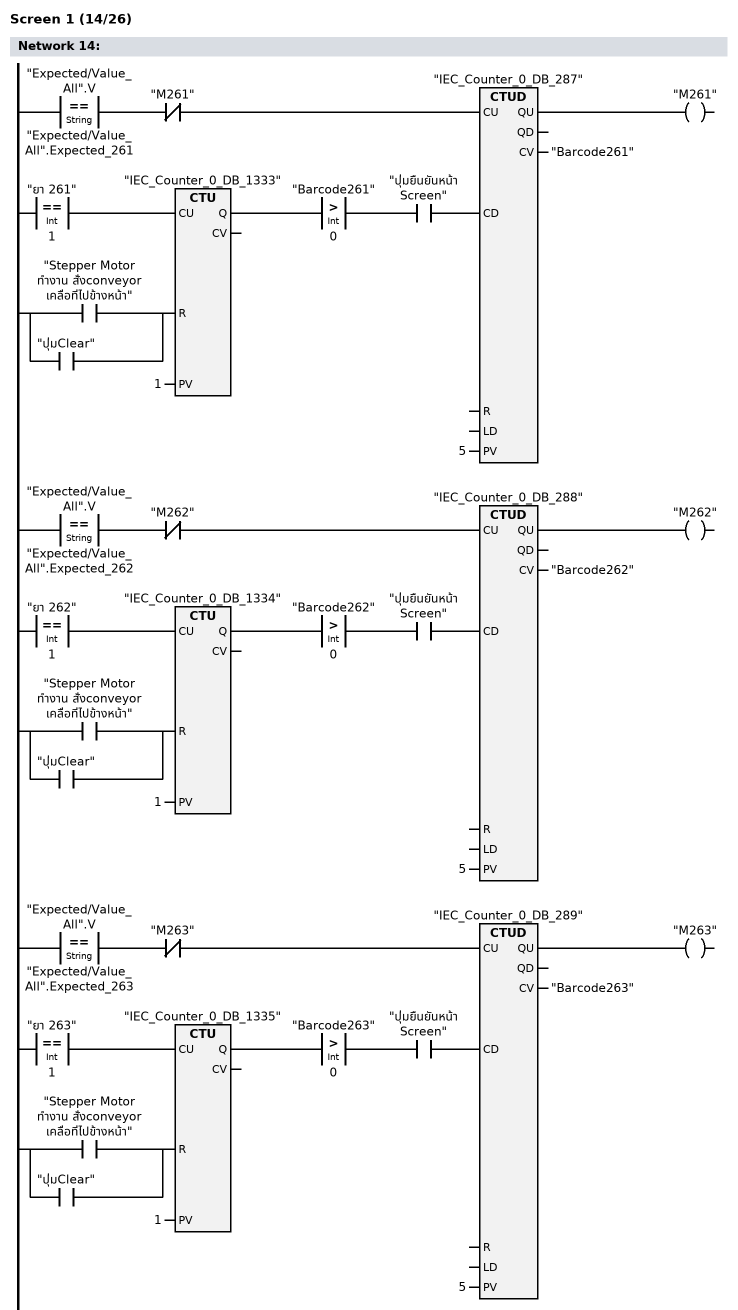
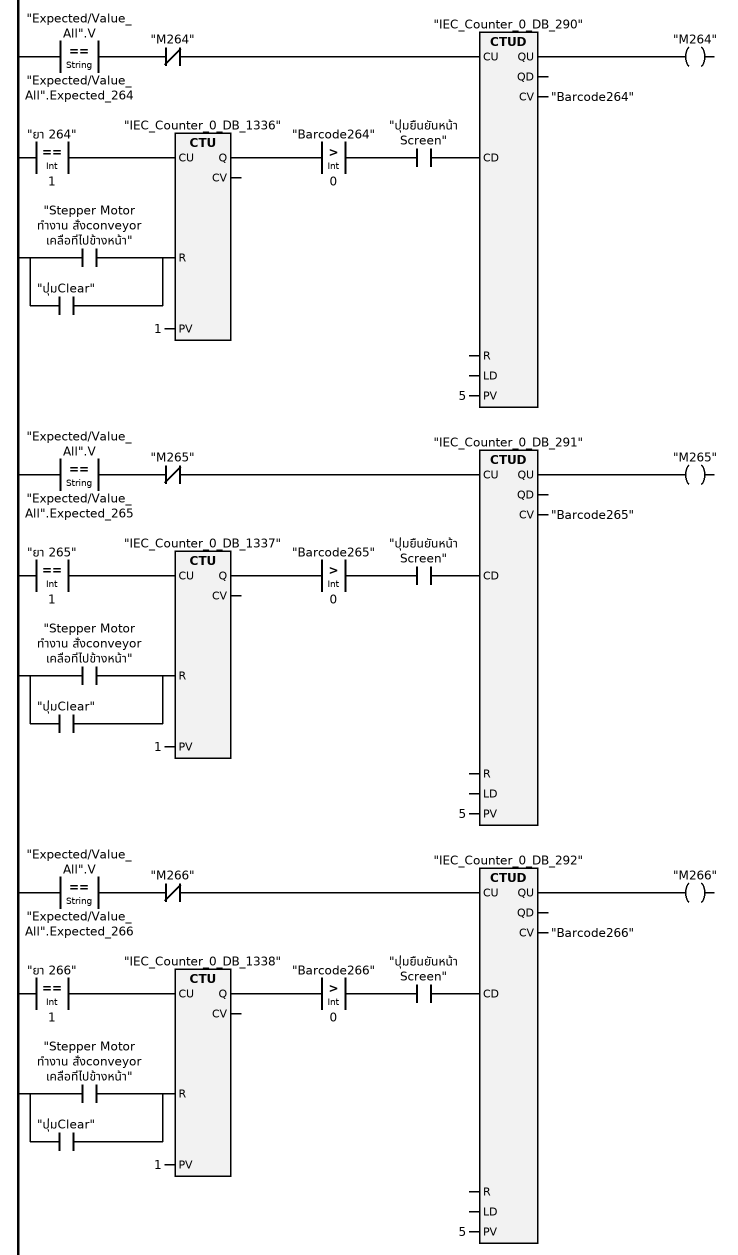
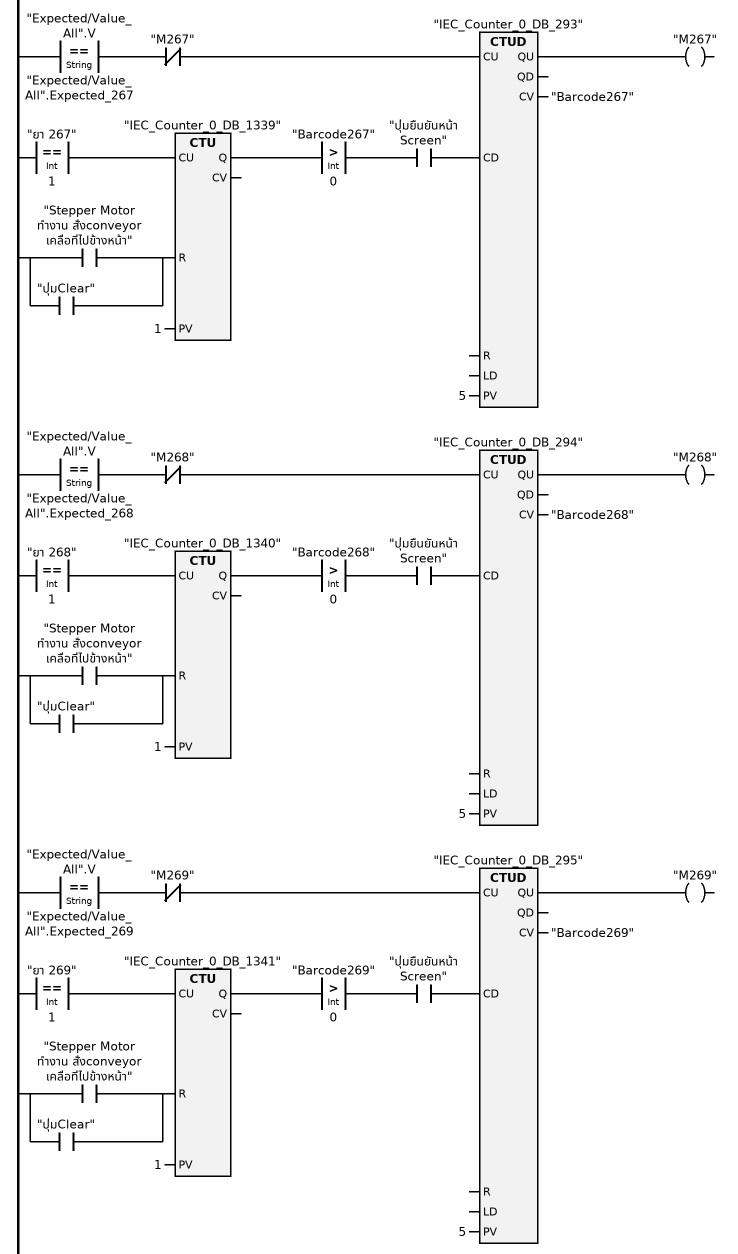
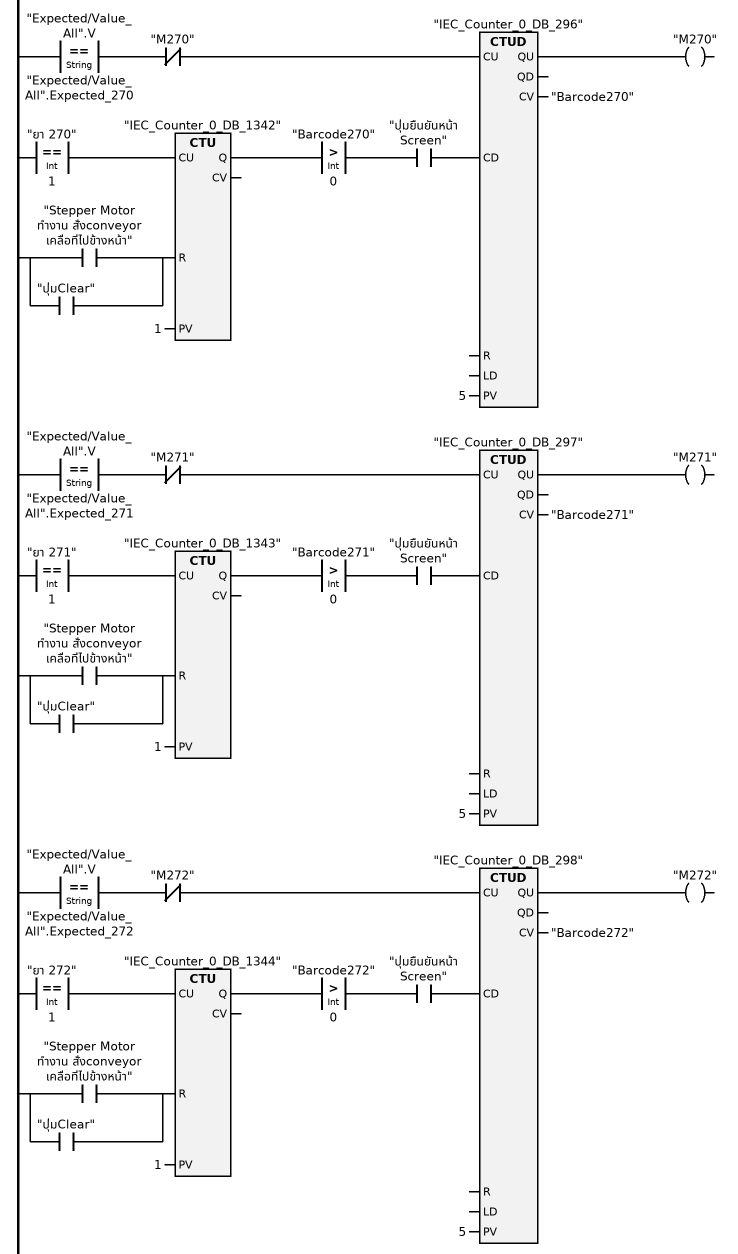
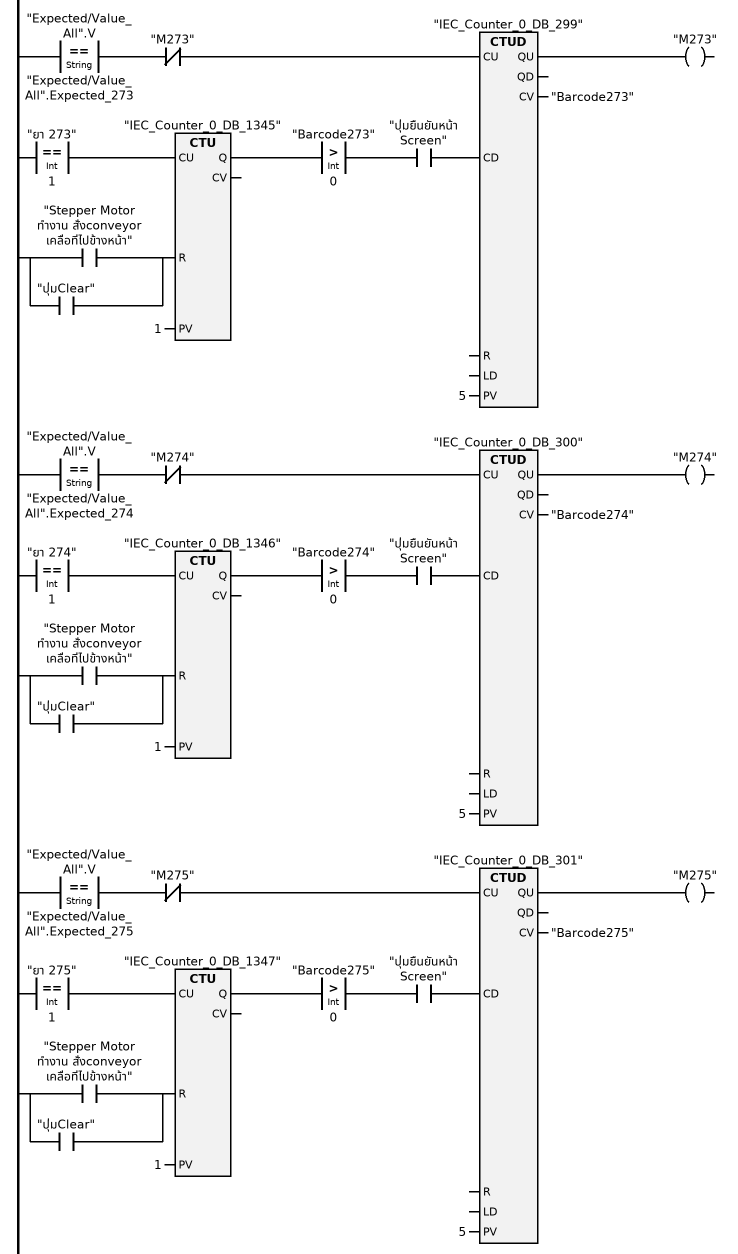
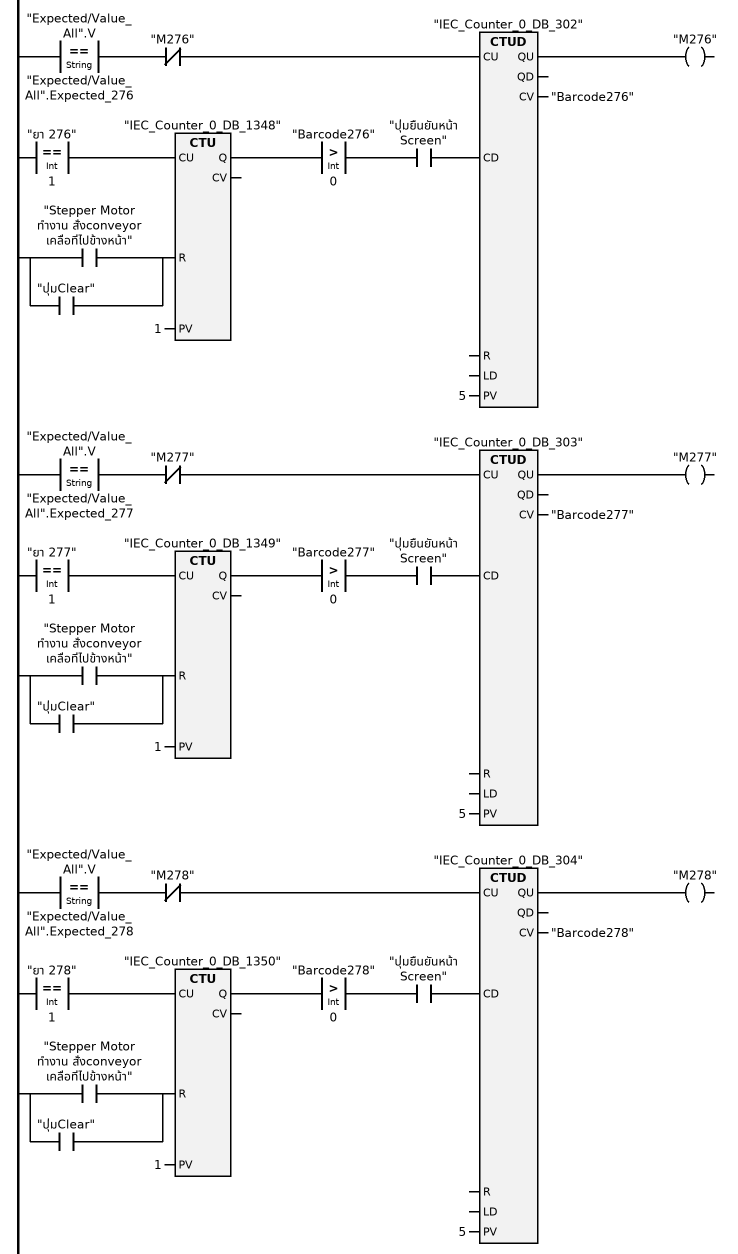
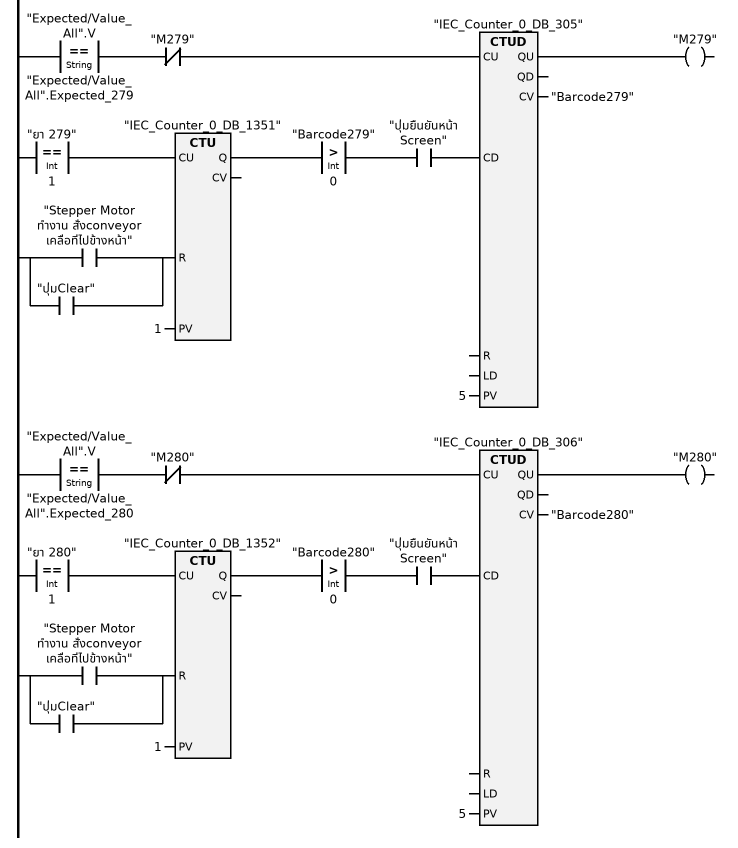
   "IEC_Counter_0_DB_1333".CTU(CU := "ยา 261" = 1,
                           R := "Stepper Motor ทำงาน สั่งconveyor เคลื่อที่ไปข้างหน้า" OR "ปุ่มClear",
                           PV := 1);
   "IEC_Counter_0_DB_287".CTUD(CU := ("Expected/Value_All".V = "Expected/Value_All".Expected_261) AND NOT "M261",
                           CD := "IEC_Counter_0_DB_1333".Q AND ("Barcode261" > 0) AND "ปุ่มยืนยันหน้า Screen",
                           PV := 5,
                           CV => "Barcode261");
   "M261" := "IEC_Counter_0_DB_287".QU;
   "IEC_Counter_0_DB_1334".CTU(CU := "ยา 262" = 1,
                           R := "Stepper Motor ทำงาน สั่งconveyor เคลื่อที่ไปข้างหน้า" OR "ปุ่มClear",
                           PV := 1);
   "IEC_Counter_0_DB_288".CTUD(CU := ("Expected/Value_All".V = "Expected/Value_All".Expected_262) AND NOT "M262",
                           CD := "IEC_Counter_0_DB_1334".Q AND ("Barcode262" > 0) AND "ปุ่มยืนยันหน้า Screen",
                           PV := 5,
                           CV => "Barcode262");
   "M262" := "IEC_Counter_0_DB_288".QU;
   "IEC_Counter_0_DB_1335".CTU(CU := "ยา 263" = 1,
                           R := "Stepper Motor ทำงาน สั่งconveyor เคลื่อที่ไปข้างหน้า" OR "ปุ่มClear",
                           PV := 1);
   "IEC_Counter_0_DB_289".CTUD(CU := ("Expected/Value_All".V = "Expected/Value_All".Expected_263) AND NOT "M263",
                           CD := "IEC_Counter_0_DB_1335".Q AND ("Barcode263" > 0) AND "ปุ่มยืนยันหน้า Screen",
                           PV := 5,
                           CV => "Barcode263");
   "M263" := "IEC_Counter_0_DB_289".QU;
   "IEC_Counter_0_DB_1336".CTU(CU := "ยา 264" = 1,
                           R := "Stepper Motor ทำงาน สั่งconveyor เคลื่อที่ไปข้างหน้า" OR "ปุ่มClear",
                           PV := 1);
   "IEC_Counter_0_DB_290".CTUD(CU := ("Expected/Value_All".V = "Expected/Value_All".Expected_264) AND NOT "M264",
                           CD := "IEC_Counter_0_DB_1336".Q AND ("Barcode264" > 0) AND "ปุ่มยืนยันหน้า Screen",
                           PV := 5,
                           CV => "Barcode264");
   "M264" := "IEC_Counter_0_DB_290".QU;
   "IEC_Counter_0_DB_1337".CTU(CU := "ยา 265" = 1,
                           R := "Stepper Motor ทำงาน สั่งconveyor เคลื่อที่ไปข้างหน้า" OR "ปุ่มClear",
                           PV := 1);
   "IEC_Counter_0_DB_291".CTUD(CU := ("Expected/Value_All".V = "Expected/Value_All".Expected_265) AND NOT "M265",
                           CD := "IEC_Counter_0_DB_1337".Q AND ("Barcode265" > 0) AND "ปุ่มยืนยันหน้า Screen",
                           PV := 5,
                           CV => "Barcode265");
   "M265" := "IEC_Counter_0_DB_291".QU;
   "IEC_Counter_0_DB_1338".CTU(CU := "ยา 266" = 1,
                           R := "Stepper Motor ทำงาน สั่งconveyor เคลื่อที่ไปข้างหน้า" OR "ปุ่มClear",
                           PV := 1);
   "IEC_Counter_0_DB_292".CTUD(CU := ("Expected/Value_All".V = "Expected/Value_All".Expected_266) AND NOT "M266",
                           CD := "IEC_Counter_0_DB_1338".Q AND ("Barcode266" > 0) AND "ปุ่มยืนยันหน้า Screen",
                           PV := 5,
                           CV => "Barcode266");
   "M266" := "IEC_Counter_0_DB_292".QU;
   "IEC_Counter_0_DB_1339".CTU(CU := "ยา 267" = 1,
                           R := "Stepper Motor ทำงาน สั่งconveyor เคลื่อที่ไปข้างหน้า" OR "ปุ่มClear",
                           PV := 1);
   "IEC_Counter_0_DB_293".CTUD(CU := ("Expected/Value_All".V = "Expected/Value_All".Expected_267) AND NOT "M267",
                           CD := "IEC_Counter_0_DB_1339".Q AND ("Barcode267" > 0) AND "ปุ่มยืนยันหน้า Screen",
                           PV := 5,
                           CV => "Barcode267");
   "M267" := "IEC_Counter_0_DB_293".QU;
   "IEC_Counter_0_DB_1340".CTU(CU := "ยา 268" = 1,
                           R := "Stepper Motor ทำงาน สั่งconveyor เคลื่อที่ไปข้างหน้า" OR "ปุ่มClear",
                           PV := 1);
   "IEC_Counter_0_DB_294".CTUD(CU := ("Expected/Value_All".V = "Expected/Value_All".Expected_268) AND NOT "M268",
                           CD := "IEC_Counter_0_DB_1340".Q AND ("Barcode268" > 0) AND "ปุ่มยืนยันหน้า Screen",
                           PV := 5,
                           CV => "Barcode268");
   "M268" := "IEC_Counter_0_DB_294".QU;
   "IEC_Counter_0_DB_1341".CTU(CU := "ยา 269" = 1,
                           R := "Stepper Motor ทำงาน สั่งconveyor เคลื่อที่ไปข้างหน้า" OR "ปุ่มClear",
                           PV := 1);
   "IEC_Counter_0_DB_295".CTUD(CU := ("Expected/Value_All".V = "Expected/Value_All".Expected_269) AND NOT "M269",
                           CD := "IEC_Counter_0_DB_1341".Q AND ("Barcode269" > 0) AND "ปุ่มยืนยันหน้า Screen",
                           PV := 5,
                           CV => "Barcode269");
   "M269" := "IEC_Counter_0_DB_295".QU;
   "IEC_Counter_0_DB_1342".CTU(CU := "ยา 270" = 1,
                           R := "Stepper Motor ทำงาน สั่งconveyor เคลื่อที่ไปข้างหน้า" OR "ปุ่มClear",
                           PV := 1);
   "IEC_Counter_0_DB_296".CTUD(CU := ("Expected/Value_All".V = "Expected/Value_All".Expected_270) AND NOT "M270",
                           CD := "IEC_Counter_0_DB_1342".Q AND ("Barcode270" > 0) AND "ปุ่มยืนยันหน้า Screen",
                           PV := 5,
                           CV => "Barcode270");
   "M270" := "IEC_Counter_0_DB_296".QU;
   "IEC_Counter_0_DB_1343".CTU(CU := "ยา 271" = 1,
                           R := "Stepper Motor ทำงาน สั่งconveyor เคลื่อที่ไปข้างหน้า" OR "ปุ่มClear",
                           PV := 1);
   "IEC_Counter_0_DB_297".CTUD(CU := ("Expected/Value_All".V = "Expected/Value_All".Expected_271) AND NOT "M271",
                           CD := "IEC_Counter_0_DB_1343".Q AND ("Barcode271" > 0) AND "ปุ่มยืนยันหน้า Screen",
                           PV := 5,
                           CV => "Barcode271");
   "M271" := "IEC_Counter_0_DB_297".QU;
   "IEC_Counter_0_DB_1344".CTU(CU := "ยา 272" = 1,
                           R := "Stepper Motor ทำงาน สั่งconveyor เคลื่อที่ไปข้างหน้า" OR "ปุ่มClear",
                           PV := 1);
   "IEC_Counter_0_DB_298".CTUD(CU := ("Expected/Value_All".V = "Expected/Value_All".Expected_272) AND NOT "M272",
                           CD := "IEC_Counter_0_DB_1344".Q AND ("Barcode272" > 0) AND "ปุ่มยืนยันหน้า Screen",
                           PV := 5,
                           CV => "Barcode272");
   "M272" := "IEC_Counter_0_DB_298".QU;
   "IEC_Counter_0_DB_1345".CTU(CU := "ยา 273" = 1,
                           R := "Stepper Motor ทำงาน สั่งconveyor เคลื่อที่ไปข้างหน้า" OR "ปุ่มClear",
                           PV := 1);
   "IEC_Counter_0_DB_299".CTUD(CU := ("Expected/Value_All".V = "Expected/Value_All".Expected_273) AND NOT "M273",
                           CD := "IEC_Counter_0_DB_1345".Q AND ("Barcode273" > 0) AND "ปุ่มยืนยันหน้า Screen",
                           PV := 5,
                           CV => "Barcode273");
   "M273" := "IEC_Counter_0_DB_299".QU;
   "IEC_Counter_0_DB_1346".CTU(CU := "ยา 274" = 1,
                           R := "Stepper Motor ทำงาน สั่งconveyor เคลื่อที่ไปข้างหน้า" OR "ปุ่มClear",
                           PV := 1);
   "IEC_Counter_0_DB_300".CTUD(CU := ("Expected/Value_All".V = "Expected/Value_All".Expected_274) AND NOT "M274",
                           CD := "IEC_Counter_0_DB_1346".Q AND ("Barcode274" > 0) AND "ปุ่มยืนยันหน้า Screen",
                           PV := 5,
                           CV => "Barcode274");
   "M274" := "IEC_Counter_0_DB_300".QU;
   "IEC_Counter_0_DB_1347".CTU(CU := "ยา 275" = 1,
                           R := "Stepper Motor ทำงาน สั่งconveyor เคลื่อที่ไปข้างหน้า" OR "ปุ่มClear",
                           PV := 1);
   "IEC_Counter_0_DB_301".CTUD(CU := ("Expected/Value_All".V = "Expected/Value_All".Expected_275) AND NOT "M275",
                           CD := "IEC_Counter_0_DB_1347".Q AND ("Barcode275" > 0) AND "ปุ่มยืนยันหน้า Screen",
                           PV := 5,
                           CV => "Barcode275");
   "M275" := "IEC_Counter_0_DB_301".QU;
   "IEC_Counter_0_DB_1348".CTU(CU := "ยา 276" = 1,
                           R := "Stepper Motor ทำงาน สั่งconveyor เคลื่อที่ไปข้างหน้า" OR "ปุ่มClear",
                           PV := 1);
   "IEC_Counter_0_DB_302".CTUD(CU := ("Expected/Value_All".V = "Expected/Value_All".Expected_276) AND NOT "M276",
                           CD := "IEC_Counter_0_DB_1348".Q AND ("Barcode276" > 0) AND "ปุ่มยืนยันหน้า Screen",
                           PV := 5,
                           CV => "Barcode276");
   "M276" := "IEC_Counter_0_DB_302".QU;
   "IEC_Counter_0_DB_1349".CTU(CU := "ยา 277" = 1,
                           R := "Stepper Motor ทำงาน สั่งconveyor เคลื่อที่ไปข้างหน้า" OR "ปุ่มClear",
                           PV := 1);
   "IEC_Counter_0_DB_303".CTUD(CU := ("Expected/Value_All".V = "Expected/Value_All".Expected_277) AND NOT "M277",
                           CD := "IEC_Counter_0_DB_1349".Q AND ("Barcode277" > 0) AND "ปุ่มยืนยันหน้า Screen",
                           PV := 5,
                           CV => "Barcode277");
   "M277" := "IEC_Counter_0_DB_303".QU;
   "IEC_Counter_0_DB_1350".CTU(CU := "ยา 278" = 1,
                           R := "Stepper Motor ทำงาน สั่งconveyor เคลื่อที่ไปข้างหน้า" OR "ปุ่มClear",
                           PV := 1);
   "IEC_Counter_0_DB_304".CTUD(CU := ("Expected/Value_All".V = "Expected/Value_All".Expected_278) AND NOT "M278",
                           CD := "IEC_Counter_0_DB_1350".Q AND ("Barcode278" > 0) AND "ปุ่มยืนยันหน้า Screen",
                           PV := 5,
                           CV => "Barcode278");
   "M278" := "IEC_Counter_0_DB_304".QU;
   "IEC_Counter_0_DB_1351".CTU(CU := "ยา 279" = 1,
                           R := "Stepper Motor ทำงาน สั่งconveyor เคลื่อที่ไปข้างหน้า" OR "ปุ่มClear",
                           PV := 1);
   "IEC_Counter_0_DB_305".CTUD(CU := ("Expected/Value_All".V = "Expected/Value_All".Expected_279) AND NOT "M279",
                           CD := "IEC_Counter_0_DB_1351".Q AND ("Barcode279" > 0) AND "ปุ่มยืนยันหน้า Screen",
                           PV := 5,
                           CV => "Barcode279");
   "M279" := "IEC_Counter_0_DB_305".QU;
   "IEC_Counter_0_DB_1352".CTU(CU := "ยา 280" = 1,
                           R := "Stepper Motor ทำงาน สั่งconveyor เคลื่อที่ไปข้างหน้า" OR "ปุ่มClear",
                           PV := 1);
   "IEC_Counter_0_DB_306".CTUD(CU := ("Expected/Value_All".V = "Expected/Value_All".Expected_280) AND NOT "M280",
                           CD := "IEC_Counter_0_DB_1352".Q AND ("Barcode280" > 0) AND "ปุ่มยืนยันหน้า Screen",
                           PV := 5,
                           CV => "Barcode280");
   "M280" := "IEC_Counter_0_DB_306".QU;
END_REGION

REGION Network 15
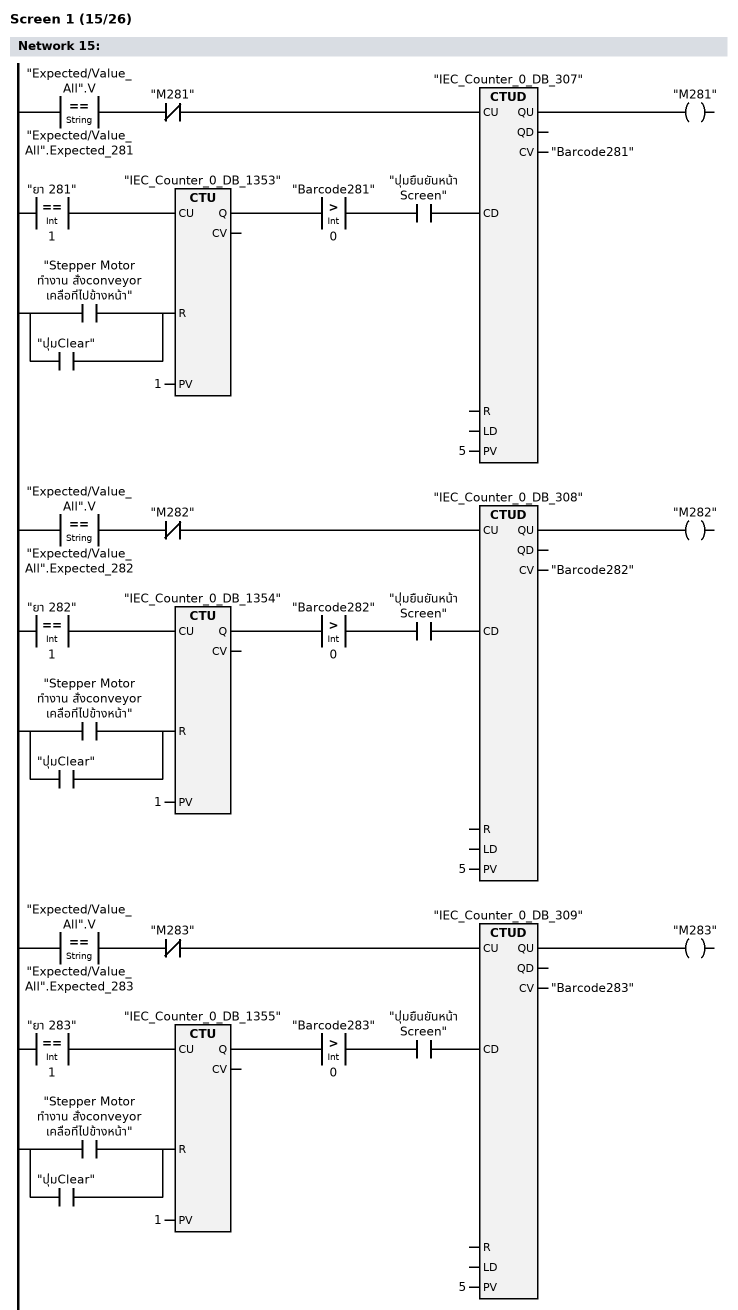
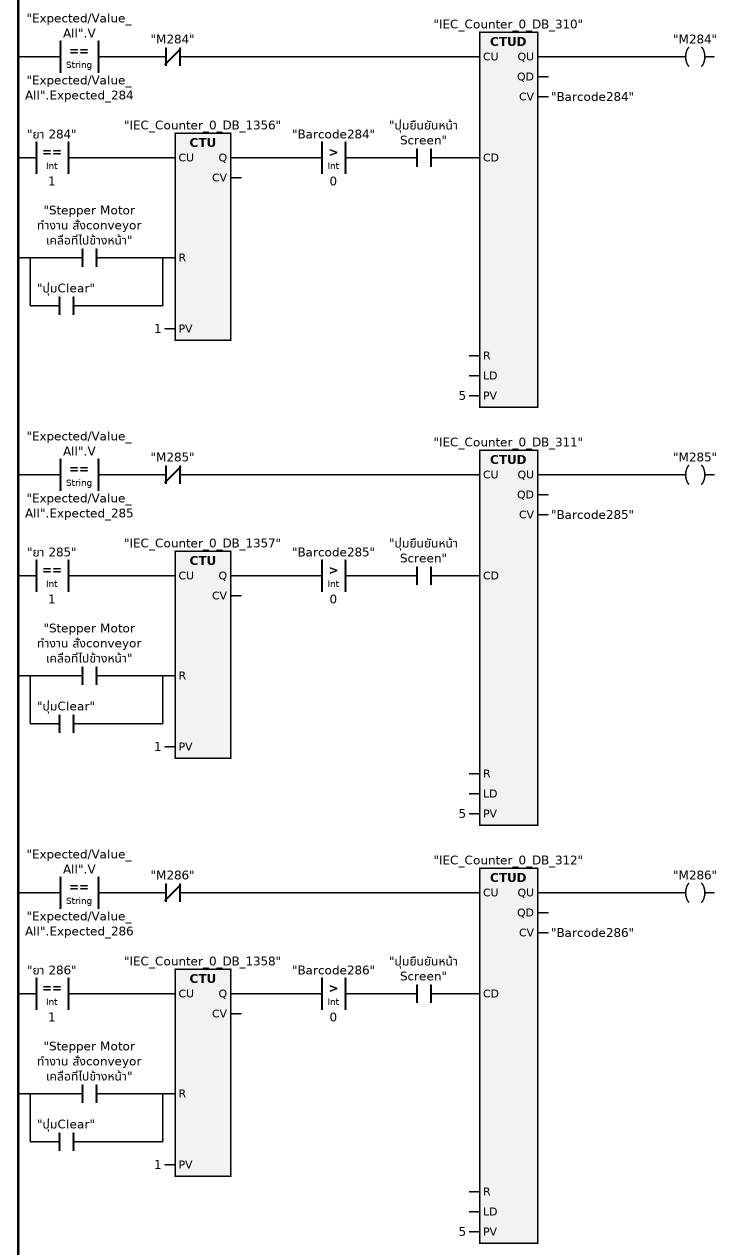
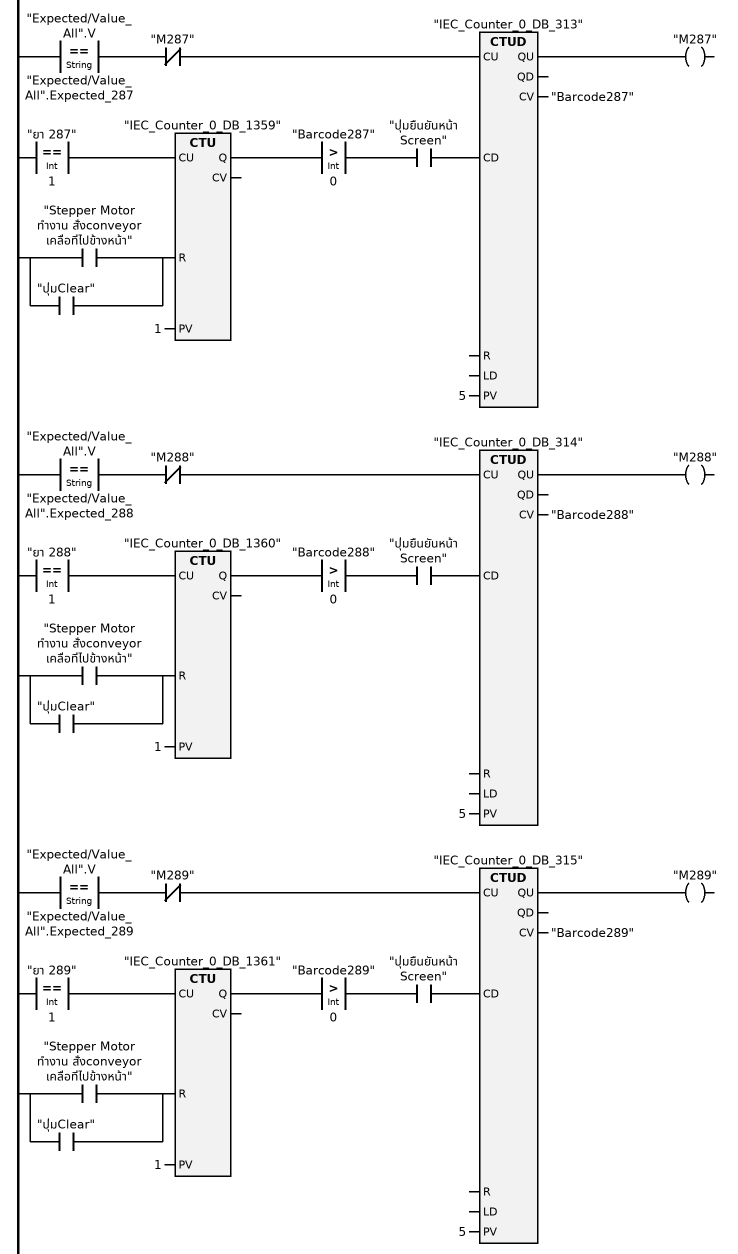
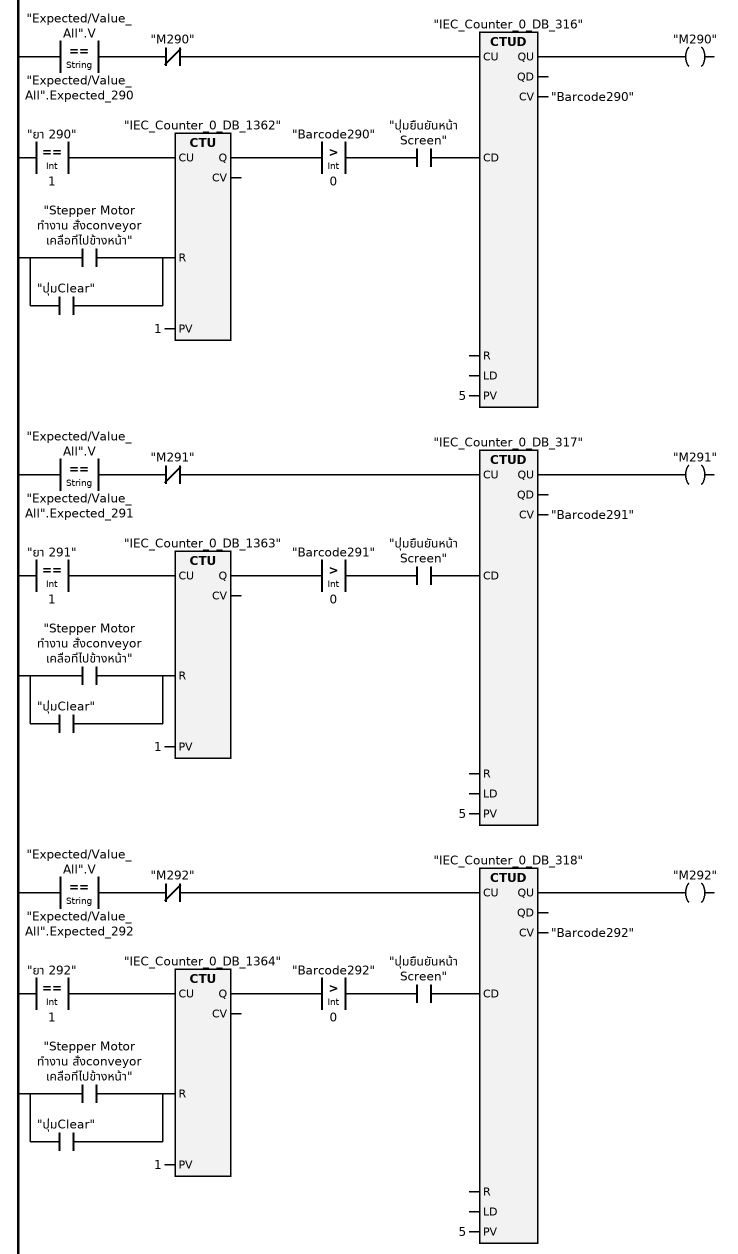
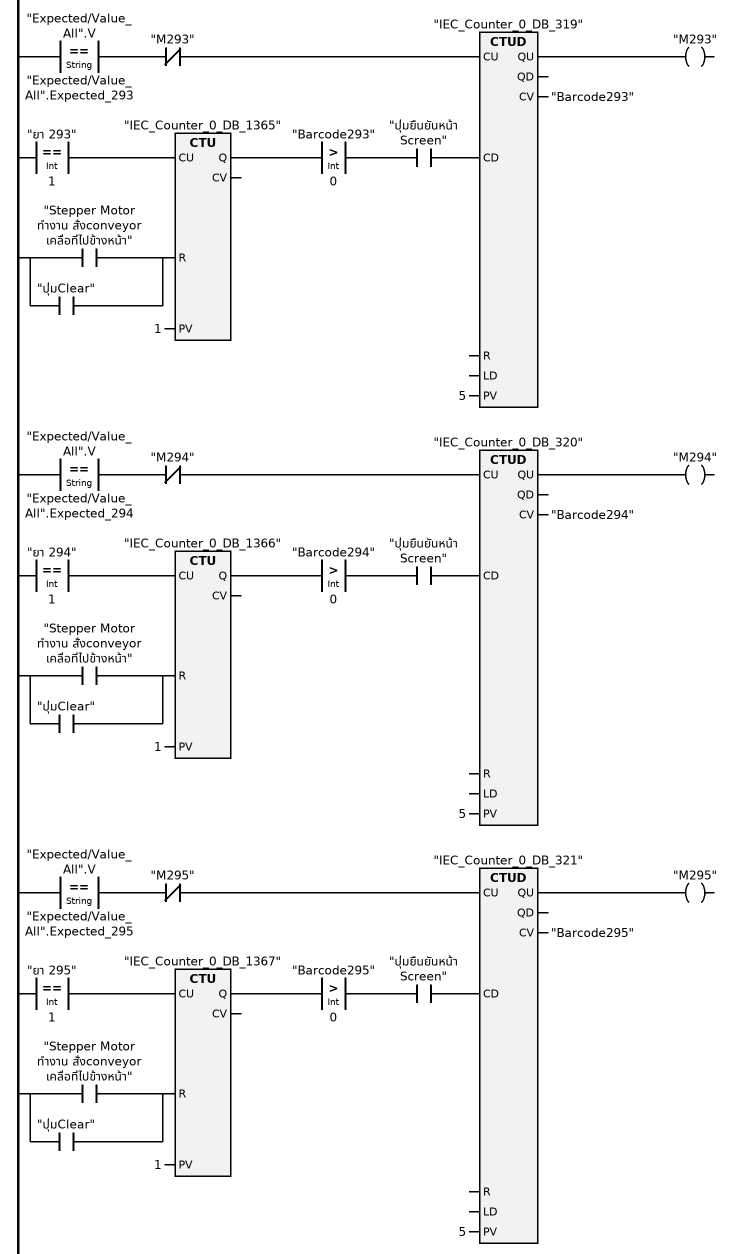
